// TIA Portal V15.1 export
ORGANIZATION_BLOCK "Startup"   // OB100, LAD, Startup
TITLE = Startup
{ S7_Optimized_Access := 'TRUE' }
VERSION : 0.1
// Startup OB (decisions/0006)
// stored: AutoNumber false, IsIECCheckEnabled false, SetENOAutomatically False
   VAR_INPUT
      LostRetentive : Bool;
      LostRTC : Bool;
   END_VAR
BEGIN

REGION Network 1: C02 — power-up: first-scan flag (scrubber trips, burners need START)
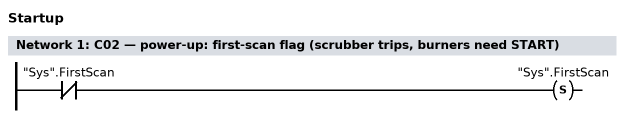
   RUNG wire#powerrail
      I_Contact( "Sys".FirstScan )
      S_Coil( "Sys".FirstScan )
   END_RUNG
   // the same network as SCL:
   IF NOT "Sys".FirstScan THEN "Sys".FirstScan := TRUE; END_IF;
END_REGION
END_ORGANIZATION_BLOCK
